(* Blister Pack Counter to Target *)

PROGRAM main
  VAR
    PillSensor AT %IX0.3 : BOOL;
    Reset AT %IX0.1 : BOOL;
    Packager AT %QX0.0 : BOOL;
    CycleComplete AT %QX0.2 : BOOL;
    Counter : INT; (* Pill Count Variable for SCADA *)
    CTU0 : CTU;
    TOF0 : TOF;
  END_VAR
  VAR  (* added by the conversion: wires and edge detectors of the diagram *)
    R_TRIG1 : R_TRIG;
  END_VAR

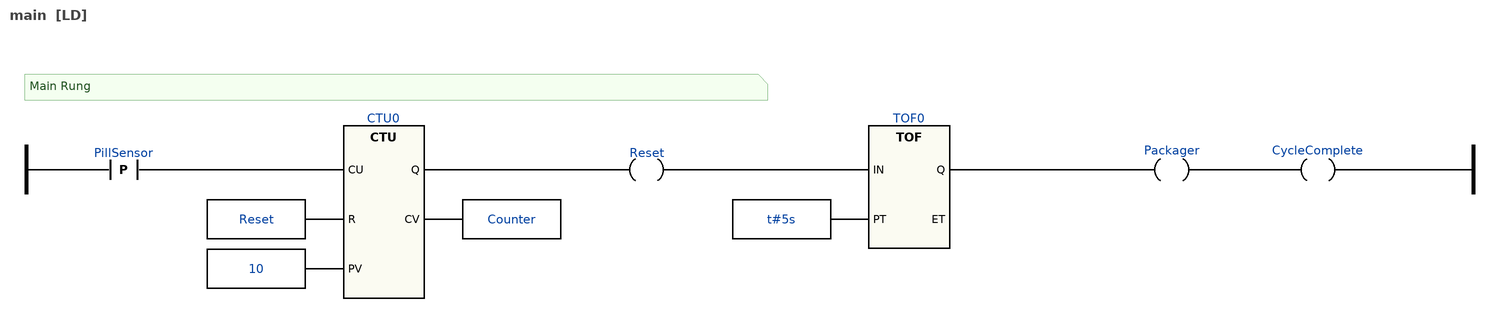
(* LD diagram, written out as Structured Text *)
(* Main Rung *)
R_TRIG1(CLK := PillSensor);
CTU0(CU := R_TRIG1.Q, R := Reset, PV := 10);
Reset := CTU0.Q;
TOF0(IN := CTU0.Q, PT := t#5s);
Packager := TOF0.Q;
CycleComplete := TOF0.Q;
Counter := CTU0.CV;
END_PROGRAM
